# B&R Automation Studio project lab1_meh1
Automation Studio 4.5.2.102

## Configuration Config1

CPU 4PP065.0571-P74, AutomationRuntime D4.52, Build 4.1.2, Vc V4.52.0

### Task classes (Cpu.sw)
```
Cyclic#1:
  Program <- Program.prg
Binaries: udbdef, TCData, ashwd, User, asfw, arconfig, sysconf, Role, ashwac, iomap
Libraries: Motor
```

### Hardware
```
4PP065_0571_P74 : 4PP065.0571-P74 v1.1.2.0
  Connector IF4:
    InternetAddress = 10.0.1.10
    SubnetMask = 255.255.255.0
  Connector IF5:
    ActivateDevice = 1
  ConfigurationID = labBR
  Simulation = 1
```

- Physical/Config1/4PP065_0571_P74/IoMap.iom: same as Physical/Config1/4PP065_0571_P74/Cpu.per
- Physical/Config1/4PP065_0571_P74/PvMap.vvm: same as Physical/Config1/4PP065_0571_P74/Cpu.per
## Logical view

Binary libraries used (declarations not repeated): operator, runtime, astime, AsIecCon


### Program Logical/Program (ANSIC)

#### Cyclic.c - Cyclic code
```c
#include <bur/plctypes.h>

#ifdef _DEFAULT_INCLUDES
	#include <AsDefault.h>
#endif

void _CYCLIC ProgramCyclic(void)
{
	if (!Enable) return;
	fb_controller.e = Speed - fb_motor.w;
	FB_Regulator(&fb_controller);
	fb_motor.u = fb_controller.u;
	FB_Motor(&fb_motor);

	fb_motor2.u = Speed * fb_motor2.ke;
	FB_Motor(&fb_motor2);

	counter++;
	Speed = 50.0f * ((counter / 50) % 2);
}
```

#### Init.c - Initialization code
```c
#include <bur/plctypes.h>

#ifdef _DEFAULT_INCLUDES
	#include <AsDefault.h>
#endif

void _INIT ProgramInit(void)
{
	counter = 0;

	fb_motor.dt = 0.01f;
	fb_motor.Tm = 0.5f;
	fb_motor.ke = 0.1f;
	fb_motor.w = 0.0f;
	fb_motor.phi = 0.0f;
	fb_motor.Integrator.out = 0.0f;

	fb_motor2.dt = 0.01f;
	fb_motor2.Tm = 0.5f;
	fb_motor2.ke = 0.1f;
	fb_motor2.w = 0.0f;
	fb_motor2.phi = 0.0f;
	fb_motor2.Integrator.out = 0.0f;

	float Tj = 0.15f;
	fb_controller.dt = 0.01f;
	fb_controller.iyOld = 0.0f;
	fb_controller.max_abs_value = 200.0f;
	fb_controller.k_p = fb_motor.ke * fb_motor.Tm / Tj;
	fb_controller.k_i = fb_motor.ke / Tj;
	fb_controller.integrator.out = 0.0f;

	Speed = 0.0f;
	Enable = 1;
}
```

#### Exit.c - Exit code
```c
#include <bur/plctypes.h>

#ifdef _DEFAULT_INCLUDES
	#include <AsDefault.h>
#endif

void _EXIT ProgramExit(void)
{

}
```

#### Variables.var - Local variables
```iecst
VAR
	fb_controller : FB_Regulator;
	fb_motor : FB_Motor;
	fb_motor2 : FB_Motor;
	counter : UDINT;
	Speed : REAL;
	Enable : BOOL;
END_VAR
```

### Library Logical/Motor (ANSIC)

#### Motor.fun - Exported functions and function blocks
```iecst
{REDUND_ERROR} {REDUND_UNREPLICABLE} FUNCTION_BLOCK FB_Integrator (*TODO: Add your comment here*) (*$GROUP=User,$CAT=User,$GROUPICON=User.png,$CATICON=User.png*)
	VAR_INPUT
		in : {REDUND_UNREPLICABLE} REAL;
	END_VAR
	VAR_OUTPUT
		out : {REDUND_UNREPLICABLE} REAL := 0.0;
	END_VAR
	VAR CONSTANT
		dt : REAL := 0.1;
	END_VAR
END_FUNCTION_BLOCK

{REDUND_ERROR} FUNCTION_BLOCK FB_Motor (*TODO: Add your comment here*) (*$GROUP=User,$CAT=User,$GROUPICON=User.png,$CATICON=User.png*)
	VAR_INPUT
		u : {REDUND_UNREPLICABLE} REAL;
	END_VAR
	VAR_OUTPUT
		w : REAL;
		phi : REAL;
	END_VAR
	VAR
		Integrator : FB_Integrator;
		Tm : REAL;
		ke : REAL;
	END_VAR
	VAR CONSTANT
		dt : REAL := 0.1;
	END_VAR
END_FUNCTION_BLOCK

{REDUND_ERROR} FUNCTION_BLOCK FB_Regulator (*TODO: Add your comment here*) (*$GROUP=User,$CAT=User,$GROUPICON=User.png,$CATICON=User.png*)
	VAR_INPUT
		e : {REDUND_UNREPLICABLE} REAL;
	END_VAR
	VAR_OUTPUT
		u : REAL;
	END_VAR
	VAR
		k_p : REAL;
		k_i : REAL;
		integrator : FB_Integrator;
		iyOld : REAL;
		max_abs_value : REAL;
	END_VAR
	VAR CONSTANT
		dt : REAL := 0.1;
	END_VAR
END_FUNCTION_BLOCK
```

#### FB_Integrator.c
```c
#include <bur/plctypes.h>
#ifdef __cplusplus
	extern "C"
	{
#endif
	#include "Motor.h"
#ifdef __cplusplus
	};
#endif
/* TODO: Add your comment here */
void FB_Integrator(struct FB_Integrator* inst)
{
	inst->out += inst->in * inst->dt;
}
```

#### FB_Motor.c
```c
#include <bur/plctypes.h>
#ifdef __cplusplus
	extern "C"
	{
#endif
	#include "Motor.h"
#ifdef __cplusplus
	};
#endif
/* TODO: Add your comment here */
void FB_Motor(struct FB_Motor* inst)
{
	inst->Integrator.in = (inst->u / inst->ke - inst->w) / inst->Tm;
	FB_Integrator(&inst->Integrator);
	inst->w = inst->Integrator.out;
	inst->phi += inst->w * inst->dt;
}
```

#### FB_Regulator.c
```c
#include <bur/plctypes.h>
#ifdef __cplusplus
	extern "C"
	{
#endif
	#include "Motor.h"
#ifdef __cplusplus
	};
#endif
/* TODO: Add your comment here */
#define min(a, b) (((a) < (b)) ? (a) : (b));

void FB_Regulator(struct FB_Regulator* inst)
{
	float var1 = inst->e * inst->k_p;
	var1 = min(inst->max_abs_value, var1);
	float var2 = inst->e * inst->k_i * inst->dt;
	var2 += inst->iyOld;
	inst->integrator.in = var2;
	FB_Integrator(&inst->integrator);
	var2 = inst->integrator.out;

	float sum = var1 + var2;
	inst->u =  min(inst->max_abs_value, sum);
	inst->iyOld = inst->u - sum;
}
```
